TYPE ST_Gr02HMIRef :
STRUCT
	stHMITOPLC				:ST_Gr02HMITOPLC;
	stPLCTOHMI				:ST_Gr02PLCTOHMI;
END_STRUCT
END_TYPE

(* stored: Version 1.1.0.1, ProductVersion 3.1.4024.15
   DUT ST_Gr02HMIRef: Id {29928505-e7ca-4bba-9f8b-6f11d10d0e4c} *)
